FUNCTION_BLOCK FB_LOADV
VAR_INPUT
	bEnable:BOOL;
	RemoteMachine : T_REMOTE_MACHINE;
	Variable_Type:E_DATA_TYPE;
	(*Appropriate to Variable type Value should be Used. rest of values will have no effect*)
	ValueByte:BYTE;
	ValueInteger:INT;
	ValueDouble:DINT;
	ValueReal:REAL;
	VariableNumber:BYTE;
END_VAR
VAR_OUTPUT
	bDone:BOOL;
	bBusy: BOOL;
	bError: BOOL;
END_VAR
VAR
	ESERVER: FB_ESERVER;
	eState:(IDLE,COMPOSE,EXECUTE,PARSE,SUCCESS_DONE,SUCCESS_PARSE,ABNORMAL_ANSWER,SOCKET_ERROR,SERVER_ERROR,DONE,ERROR);
	sAnswer: STRING(255);
	delimiter: ARRAY[0..100]OF UINT;
	i: UINT;
	length: UINT;
	position:UINT;
	integer: DINT;
	fraction: REAL;
END_VAR

eServer.RemoteMachine:=RemoteMachine;
eServer.eCommand:=E_COMMAND.LOADV;


CASE	eState OF
IDLE:
	bBusy:=FALSE;
	IF	bEnable	THEN
		eState:=COMPOSE;
		bDone:=FALSE;
		bBusy:=TRUE;
		bError:=FALSE;
	END_IF;
COMPOSE:
	(*	if data to be sent compose eServer.sCommandData to contain CommandData string	*)
	(*	Do not forget to strt with eServer.sCommandData:=''; to avoid send buffer repetition	*)
	eServer.sCommandData:='';
	eServer.sCommandData:=CONCAT(eServer.sCommandData,INT_TO_STRING(Variable_type));
	eServer.sCommandData:=CONCAT(eServer.sCommandData,',');
	eServer.sCommandData:=CONCAT(eServer.sCommandData,BYTE_TO_STRING(VariableNumber));
	eServer.sCommandData:=CONCAT(eServer.sCommandData,',');
	CASE Variable_Type OF
		BYTE_TYPE:
			eServer.sCommandData:=CONCAT(eServer.sCommandData,BYTE_TO_STRING(ValueByte));
		INTEGER_TYPE:
			eServer.sCommandData:=CONCAT(eServer.sCommandData,INT_TO_STRING(ValueInteger));
		DOUBLE_TYPE:
			eServer.sCommandData:=CONCAT(eServer.sCommandData,DINT_TO_STRING(ValueDouble));
		REAL_TYPE:
			eServer.sCommandData:=CONCAT(eServer.sCommandData,REAL_TO_STRING(integer+fraction));

		ROBOT_AXIS_TYPE:;
		BASE_AXIS_TYPE:;
		STATION_AXIS_TYPE:;
	END_CASE;
	eServer.sCommandData:=CONCAT(eServer.sCommandData,'$R');
	eState:=EXECUTE;
EXECUTE:
	eServer.bExecute:=TRUE;
	eServer();
	IF	eServer.bDone	THEN
		eState:=PARSE;
		eServer.bExecute:=FALSE;
		eServer();
	ELSIF	eServer.bError	THEN
		eState:=SERVER_ERROR;
		eServer.bExecute:=FALSE;
		eServer();
	END_IF;
PARSE:
	IF	eServer.sAnswer='0000$R$N' THEN
		eState:=SUCCESS_DONE;;
	ELSIF	RIGHT(eServer.sAnswer,1)='$R'	THEN
		eState:=SUCCESS_PARSE;
	ELSIF	LEFT(eServer.sAnswer,6)='ERROR: ['	THEN
		eState:=ABNORMAL_ANSWER;
	ELSE
		eState:=SOCKET_ERROR;
	END_IF;
SUCCESS_DONE:
	eState:=DONE;
SUCCESS_PARSE:
	(*
		sAnswer:=eServer.sAnswer;
		FOR i:=0 TO (SIZEOF(delimiter)/2)-1 DO
			delimiter[i]:=0;
		END_FOR;
		FOR i:=1 TO (SIZEOF(delimiter)/2)-1 DO
			delimiter[i]:=delimiter[i-1]+FIND(sAnswer,',');
			IF	delimiter[i]=delimiter[i-1]	THEN
				delimiter[i]:=delimiter[i]+FIND(sAnswer,'$R');
				EXIT;
			END_IF;
			sAnswer:=DELETE(sAnswer,delimiter[i],1);
		END_FOR;

		FOR i:=1 TO  NumberOfContactPoints/8 DO
			length:=delimiter[i]-delimiter[i-1]-1;
			position:=delimiter[i-1]+1;
			ContactPoints[i-1]:=STRING_TO_BYTE(MID(eServer.sAnswer,length,position));
		END_FOR;
*)
		eState:=DONE;
ABNORMAL_ANSWER:
	eState:=ERROR;
SOCKET_ERROR:
	eState:=ERROR;
SERVER_ERROR:
	eState:=ERROR;
DONE:
	bDone:=TRUE;
	eState:=IDLE;
ERROR:
	bError:=TRUE;
	eState:=IDLE;
END_CASE;

END_FUNCTION_BLOCK

(* stored: Version 1.1.0.1, ProductVersion 3.1.4024.16
   POU FB_LOADV: Id {66db1f28-df83-454c-8bfc-a62b8b0885ca}, SpecialFunc None *)
